(* IEC 61131-3 sources: crb-codesys/generation/scripts/repoeval/plc_hello_mixing_tank/global, 2 files *)

(* ---- HMI.st ---- *)
{attribute 'qualified_only'}
VAR_GLOBAL
	///Command to start the mixer
	MixerRunCmd: BOOL;
	///Command to stop the mixer
	MixerStopCmd: BOOL;
	///Command to open medium 1 valve
	Medium1OpenCmd: BOOL;
	///Command to close medium 1 valve
	Medium1CloseCmd: BOOL;
	///Command to open medium 2 valve
	Medium2OpenCmd: BOOL;
	///Command to close medium 2 valve
	Medium2CloseCmd: BOOL;
	///Command to open drain valve
	DrainOpenCmd: BOOL;
	///Command to close drain valve
	DrainCloseCmd: BOOL;
	///Command to set the system to auto mode
	SetToAuto: BOOL;
	///Command to set the system to manual mode
	SetToManual: BOOL;
	//HMI Support variables
	MotorRotating : REAL;
	//System in AUTO
	InAuto : BOOL;
	//System in MANUAL
	InManual : BOOL;
	//Cycles completed
	CyclesCompleted : UINT;
END_VAR

(* ---- IO.st ---- *)
{attribute 'qualified_only' := ''}
VAR_GLOBAL
	///Tank level switch (HIGH) active
	xDI_LS01_TankLevelFull: BOOL;
	///Tank level switch (LOW) active
	xDI_LS02_TankLevelEmpty: BOOL;
	///Medium 1 filling valve open
	xDI_VV01_Medium1_Opened: BOOL;
	///Medium 2 filling valve open
	xDI_VV02_Medium2_Opened: BOOL;
	///Tank draining valve open
	xDI_VV03_TankDrain_Opened: BOOL;
	///Mixer motor running
	xDI_M1_MixerMotorRunning: BOOL;
	///Medium 1 filling valve open command
	xDO_VV01_Medium1_OpenCmd: BOOL;
	///Medium 2 filling valve open command
	xDO_VV02_Medium2_OpenCmd: BOOL;
	///Tank draining valve open command
	xDO_VV03_TankDrain_OpenCmd: BOOL;
	///Mixer motor run command
	xDO_M1_MixerMotorRunCmd: BOOL;
END_VAR
